Fanuc KAREL source: kt00261.KL

-- PROVISIONAL review KL for V770-1; original PC SHA256 03e1c0a3371b9fa24d4ae02fe0ac0d8621c25f6992db0c82e1897346be136032
-- Incomplete behavior may be omitted. Consult companion uncertainty JSON. Do not deploy.
PROGRAM KT00261
%NOLOCKGROUP
VAR
  R1 : REAL
  I2 : INTEGER
  OUT : BOOLEAN
BEGIN
  -- UNRESOLVED_PC offsets 5-16; opcodes 2E,23
  -- UNRESOLVED_PC offsets 21-32; opcodes 2E,23
  -- UNRESOLVED_PC offsets 37-57; opcodes 21,21,64,6D,23
  -- UNRESOLVED_PC offsets 62-66; opcodes 7F
END KT00261
